(* IEC 61131-3 sources: Test-Git_ESME26/TestProgettoESME_26.fbsproj/PacDriveLib Migration/Motion/Control/Brake/FB_BrakeCouplingTime.fb.st^, 4 files *)

(* ---- ifBrake.prop.st ---- *)
PROPERTY ifBrake : DDI.IF_Brake
__SETTERDECLARATION__
VAR
END_VAR
__SETTERIMPLEMENTATION__
ifBrake_loc := ifBrake;

(* ---- Job.meth.st ---- *)
{attribute 'conditionalshow_all_locals'}
METHOD Job : BOOL

IF ifBrake_loc.BrakeCouplingTime > 0 THEN
	tBrakeCouplingTemp := DINT_TO_TIME(ifBrake_loc.BrakeCouplingTime);
ELSE
	tBrakeCouplingTemp := T#500MS;
END_IF

(* ---- timTime.prop.st ---- *)
PROPERTY INTERNAL timTime : TIME
__GETTERDECLARATION__
VAR
END_VAR
__GETTERIMPLEMENTATION__
timTime:= tBrakeCouplingTemp;

(* ---- xDone.prop.st ---- *)
PROPERTY xDone : BOOL
__SETTERDECLARATION__
VAR
END_VAR
__SETTERIMPLEMENTATION__
xDone_loc := xDone;
__GETTERDECLARATION__
VAR
END_VAR
__GETTERIMPLEMENTATION__
xDone := xDone_loc;
